(* IEC 61131-3 sources: codesys-to-s7/tests/corpus/C2S7-NAME-LEN/neg, 1 file *)

(* ---- input.st ---- *)
FUNCTION_BLOCK FB_Case
VAR
    a : INT;
END_VAR
a := 1;
END_FUNCTION_BLOCK
